(* PLC project LFAM, CODESYS CODESYS V3.5 SP22 Patch 4 *)
(* stored: creationDateTime 2026-11-11T00:00:00, modificationDateTime 2026-11-11T00:00:00 *)

PROGRAM PLC_PRG
  VAR
    PT_FUNDIDO_MPA : REAL;
    PT_FUNDIDO_RAW : INT;
    TT_SUBSTRATO_C : REAL;
    TT_SUBSTRATO_RAW : INT;
    TT_Z1 : REAL;
    TT_Z1_RAW : INT;
    TC_Z1_ABERTO : BOOL;
    TT_Z2 : REAL;
    TT_Z2_RAW : INT;
    TC_Z2_ABERTO : BOOL;
    TT_Z3 : REAL;
    TT_Z3_RAW : INT;
    TC_Z3_ABERTO : BOOL;
    TT_Z4 : REAL;
    TT_Z4_RAW : INT;
    TC_Z4_ABERTO : BOOL;
    TT_Z5 : REAL;
    TT_Z5_RAW : INT;
    TC_Z5_ABERTO : BOOL;
    TC_Z1_OK : BOOL;
    TC_Z2_OK : BOOL;
    TC_Z3_OK : BOOL;
    TC_Z4_OK : BOOL;
    TC_Z5_OK : BOOL;
    PLC_HEARTBEAT : INT;
    PWM_FASE : INT;
    PID_Z1 : Util.PID;
    SP_Z1 : REAL;
    Y_Z1 : REAL;
    LIM_Z1 : BOOL;
    OVF_Z1 : BOOL;
    PID_Z2 : Util.PID;
    SP_Z2 : REAL;
    Y_Z2 : REAL;
    LIM_Z2 : BOOL;
    OVF_Z2 : BOOL;
    PID_Z3 : Util.PID;
    SP_Z3 : REAL;
    Y_Z3 : REAL;
    LIM_Z3 : BOOL;
    OVF_Z3 : BOOL;
    PID_Z4 : Util.PID;
    SP_Z4 : REAL;
    Y_Z4 : REAL;
    LIM_Z4 : BOOL;
    OVF_Z4 : BOOL;
    PID_Z5 : Util.PID;
    SP_Z5 : REAL;
    Y_Z5 : REAL;
    LIM_Z5 : BOOL;
    OVF_Z5 : BOOL;
    PWM_Z1 : BOOL;
    PWM_Z2 : BOOL;
    PWM_Z3 : BOOL;
    PWM_Z4 : BOOL;
    PWM_Z5 : BOOL;
    PID_IR : Util.PID;
    SP_IR_C : REAL;
    Y_IR : REAL;
    LIM_IR : BOOL;
    OVF_IR : BOOL;
    PWM_IR : BOOL;
    SOBRETEMP_390_Z1 : BOOL;
    SOBRETEMP_390_Z2 : BOOL;
    SOBRETEMP_390_Z3 : BOOL;
    SOBRETEMP_390_Z4 : BOOL;
    SOBRETEMP_390_Z5 : BOOL;
    SOBRETEMP_400_Z1 : BOOL;
    SOBRETEMP_400_Z2 : BOOL;
    SOBRETEMP_400_Z3 : BOOL;
    SOBRETEMP_400_Z4 : BOOL;
    SOBRETEMP_400_Z5 : BOOL;
    SOBRETEMP_400 : BOOL;
    TC_FAULT : BOOL;
    TT_RESF : REAL;
    RESF_ACIMA_100 : BOOL;
    T_RESF_100C : TON;
    FALHA_RESF_2M : BOOL;
    EST_EXTRUSAO : BOOL;
    FUNIL_BAIXO : BOOL;
    ALIM_FUNIL : BOOL;
    T_FUNIL_VAZIO : TON;
    FALHA_SEM_MAT : BOOL;
    INV_RUN : BOOL;
    VENT_OK : BOOL;
    T_FALHA_VENT : TON;
    FALHA_VENT_10S : BOOL;
    K1_AQUEC : BOOL;
    K1_CONF : BOOL;
    T_K1_COLADO : TON;
    FALHA_K1_COL : BOOL;
    RESF_HI : BOOL;
    RESF_LO : BOOL;
    ALM_PRESSAO_16_5 : BOOL;
    PRESSAO_ALTA_17 : BOOL;
    SEG_OK : BOOL;
    MOT_SOBRETEMP : BOOL;
    INV_FALHA : BOOL;
    M_CAUSA : BOOL;
    FALHA_GERAL : BOOL;
    CAUSA_SEG_OK : BOOL;
    CAUSA_MOT_SOBRETEMP : BOOL;
    CAUSA_INV_FALHA : BOOL;
    CAUSA_PRESSAO_ALTA_17 : BOOL;
    CAUSA_SOBRETEMP_400 : BOOL;
    CAUSA_TC_FAULT : BOOL;
    CAUSA_FALHA_RESF_2M : BOOL;
    CAUSA_FALHA_SEM_MAT : BOOL;
    CAUSA_FALHA_VENT_10S : BOOL;
    CAUSA_FALHA_K1_COL : BOOL;
    BT_RESET : BOOL;
    BT_AQUEC : BOOL;
    EST_AQUEC : BOOL;
    DISJ_AQUEC : BOOL;
    RESF_ON : BOOL;
    Z1_ATEMP : BOOL;
    Z2_ATEMP : BOOL;
    Z3_ATEMP : BOOL;
    Z4_ATEMP : BOOL;
    Z5_ATEMP : BOOL;
    EST_ENCHARQUE : BOOL;
    T_ENCHARQUE : TON;
    ENCH_OK : BOOL;
    SECADOR_OK : BOOL;
    INV_PRONTO : BOOL;
    EST_PRONTO : BOOL;
    ROBO_EXT_PRONTA : BOOL;
    BT_DESLIGA : BOOL;
    SEL_AUTO : BOOL;
    BT_LIGA : BOOL;
    ROBO_CMD_EXTR : BOOL;
    VENT_MOTOR : BOOL;
    T_POS_VENT : TON;
    VENT_FIM : BOOL;
    REF_RPM_LIM : REAL;
    SP_RPM_OPERADOR : REAL;
    INV_REF : INT;
    SSR_Z1 : BOOL;
    SSR_Z2 : BOOL;
    SSR_Z3 : BOOL;
    SSR_Z4 : BOOL;
    SSR_Z5 : BOOL;
    IR_ACIMA_MIN : BOOL;
    IR_ABAIXO_MAX : BOOL;
    ROBO_EM_MOV : BOOL;
    IR_HAB : BOOL;
    SSR_IR : BOOL;
    TT_ZSR : REAL;
    ZSR_ABAIXO : BOOL;
    ALM_ZSR_BAIXA : BOOL;
    LUZ_VERDE : BOOL;
    LUZ_AMARELA : BOOL;
    LUZ_VERM_SIRENE : BOOL;
    RT_FUNIL : R_TRIG;
    FUNIL_PULSO : BOOL;
    CTU_LOTES : CTU;
    HMI_RESET_LOTES : BOOL;
    CONT_LOTES : WORD;
  END_VAR

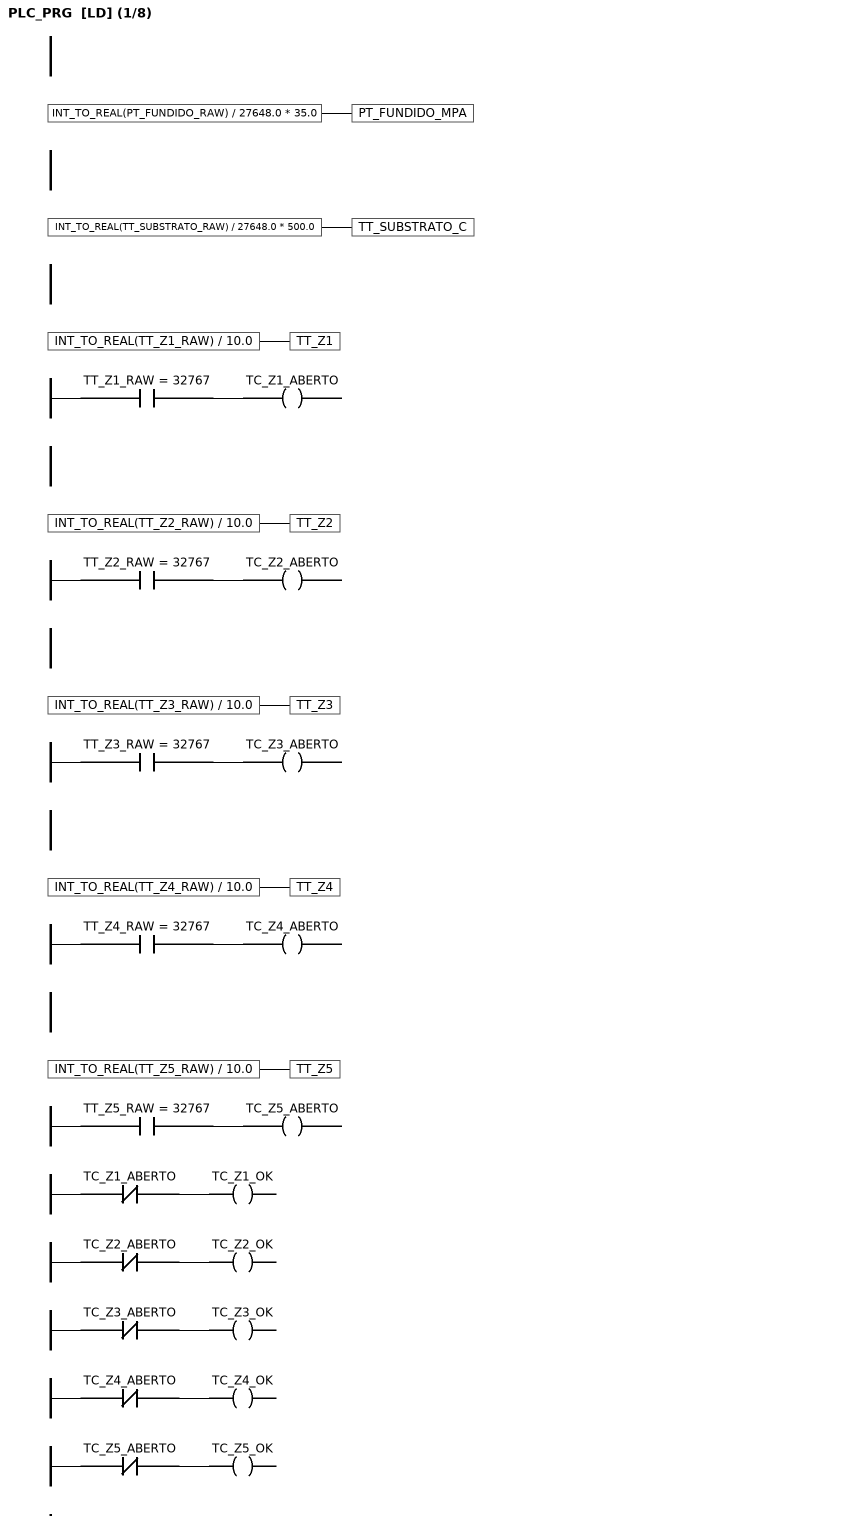
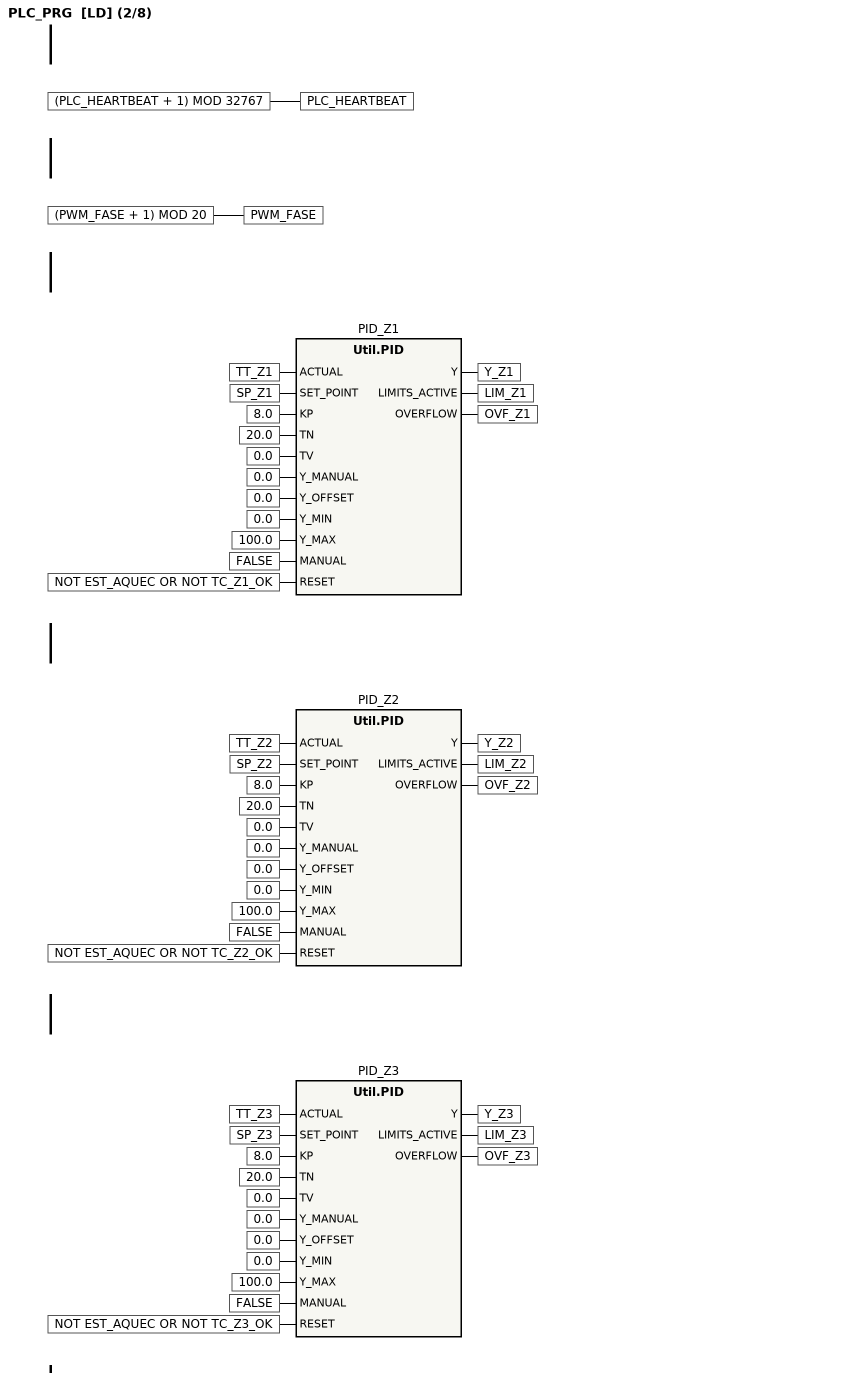
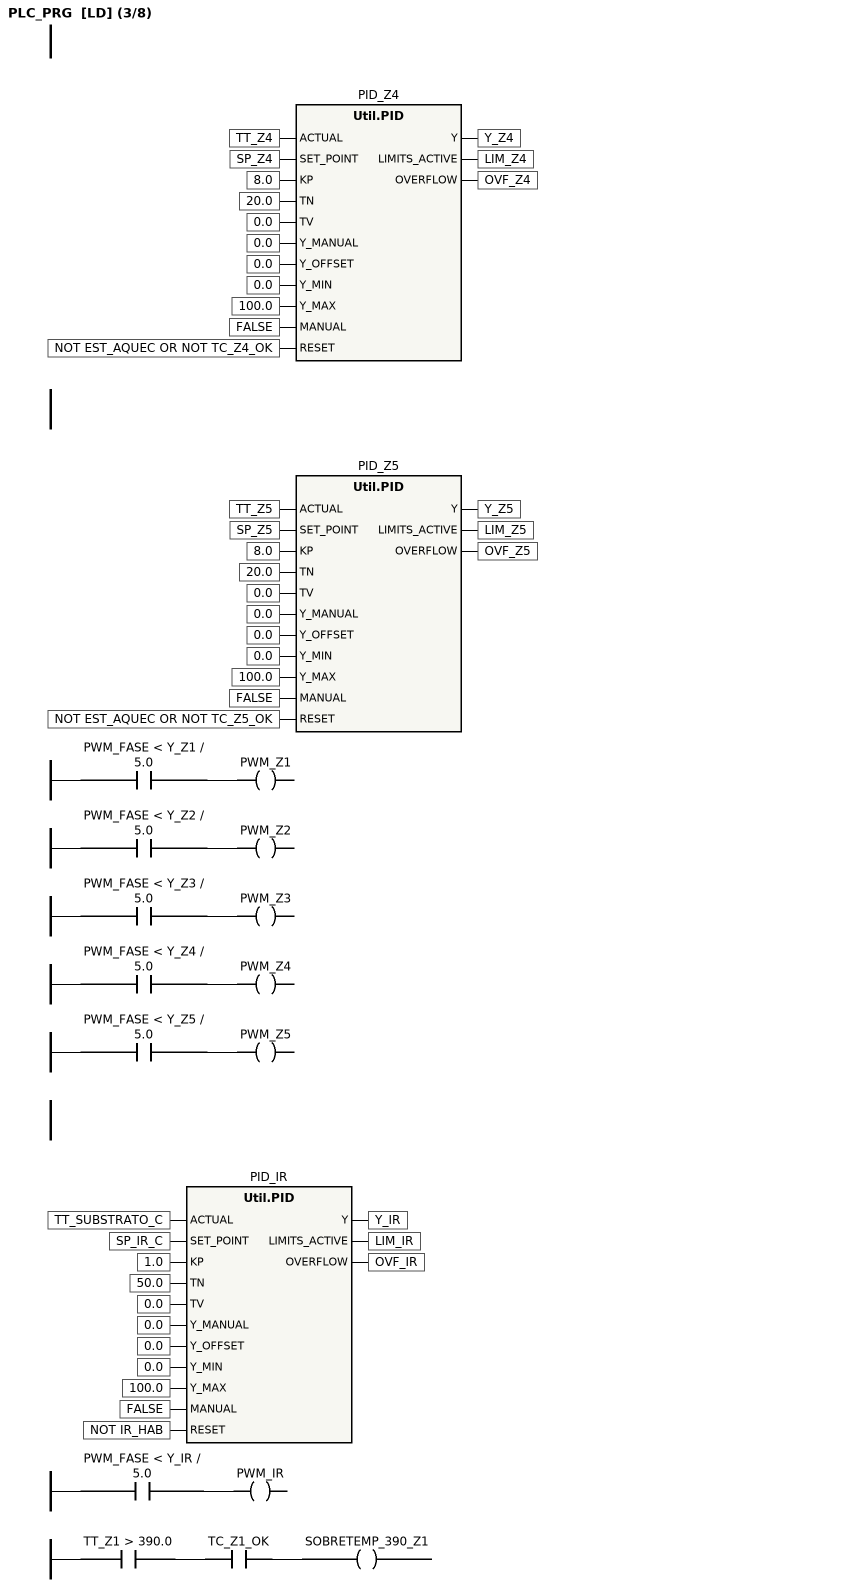
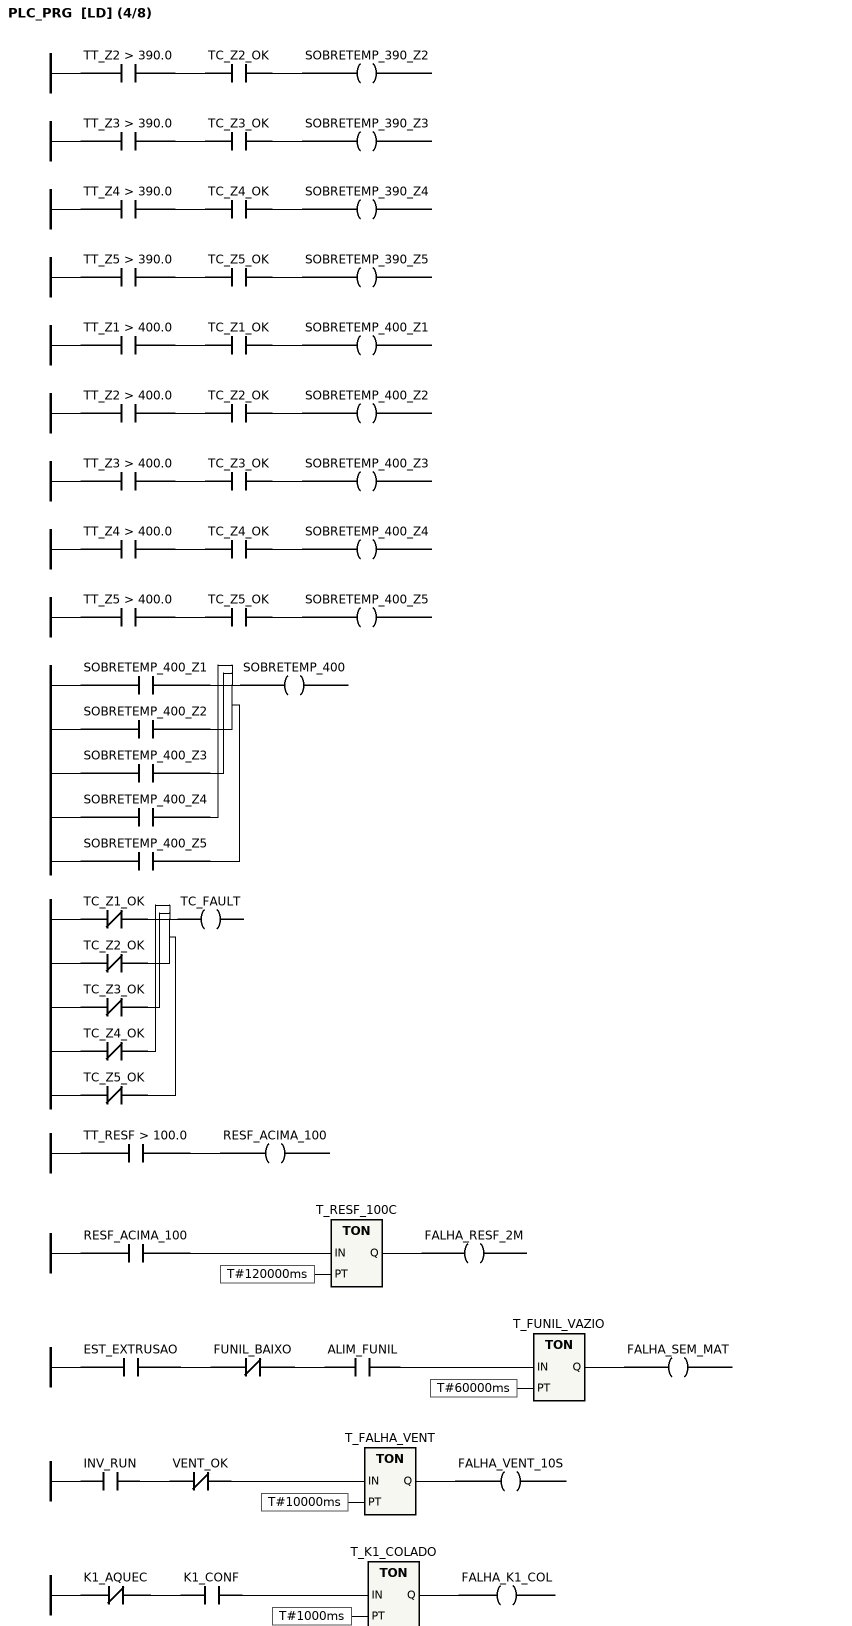
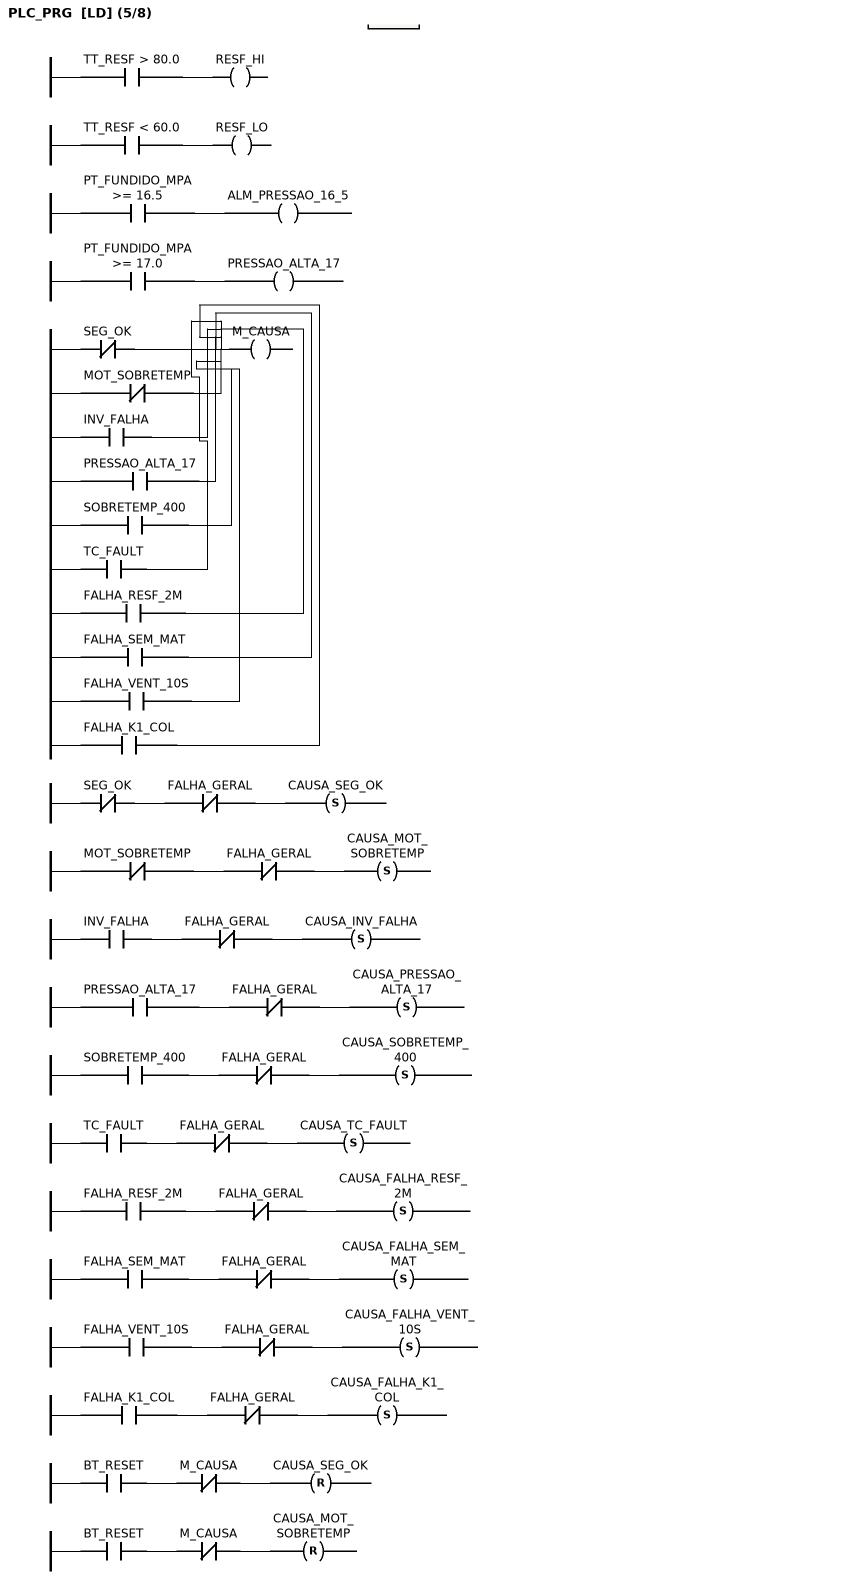
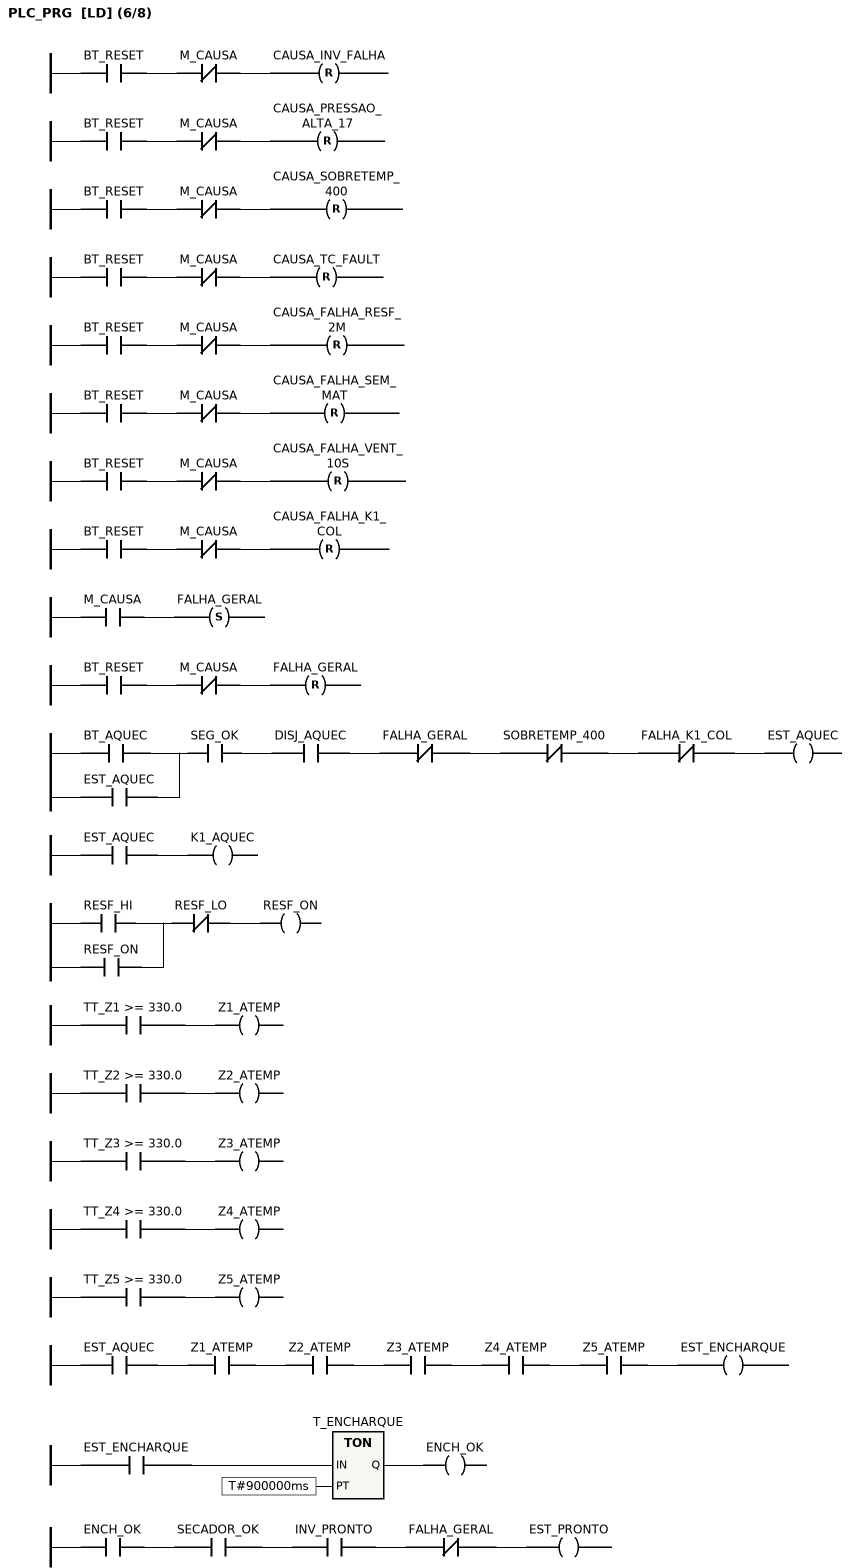
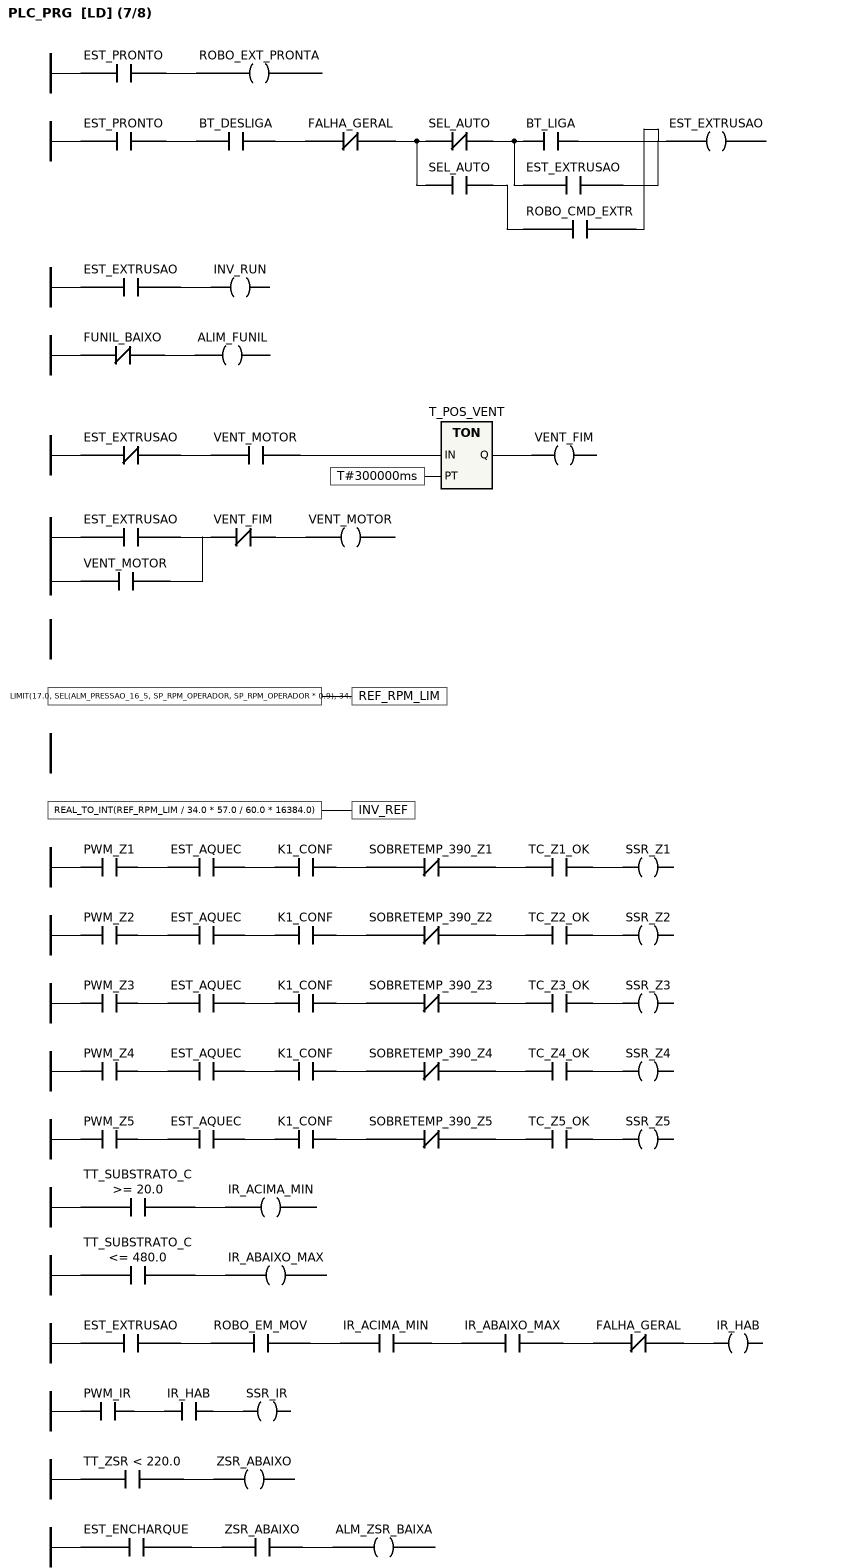
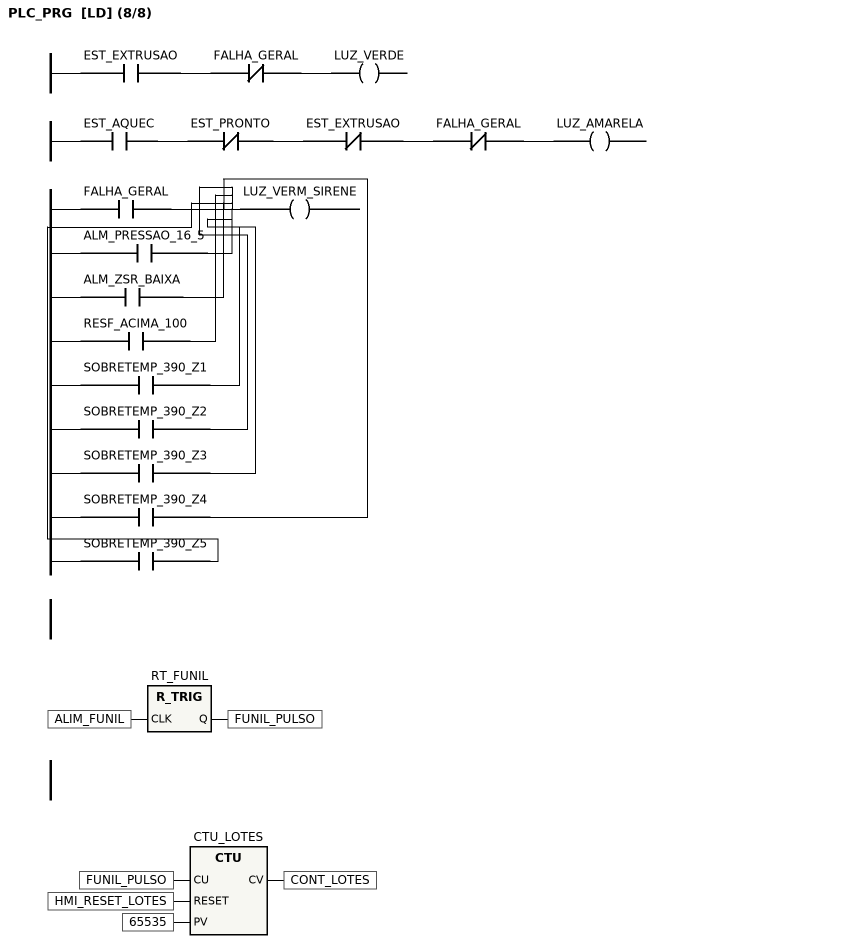
(* LD diagram, written out as Structured Text *)
(* NETWORK 01 - PT_FUNDIDO 0..27648 -> 0..35 MPa *)
PT_FUNDIDO_MPA := INT_TO_REAL(PT_FUNDIDO_RAW) / 27648.0 * 35.0;
(* NETWORK 01 - TT_SUBSTRATO 0..27648 -> 0..500 degC *)
TT_SUBSTRATO_C := INT_TO_REAL(TT_SUBSTRATO_RAW) / 27648.0 * 500.0;
(* NETWORK 02 - TT_Z1 (0,1 degC -> degC) *)
TT_Z1 := INT_TO_REAL(TT_Z1_RAW) / 10.0;
(* NETWORK 02 - Z1 termopar aberto (RAW = 32767) *)
TC_Z1_ABERTO := TT_Z1_RAW = 32767;
(* NETWORK 02 - TT_Z2 (0,1 degC -> degC) *)
TT_Z2 := INT_TO_REAL(TT_Z2_RAW) / 10.0;
(* NETWORK 02 - Z2 termopar aberto (RAW = 32767) *)
TC_Z2_ABERTO := TT_Z2_RAW = 32767;
(* NETWORK 02 - TT_Z3 (0,1 degC -> degC) *)
TT_Z3 := INT_TO_REAL(TT_Z3_RAW) / 10.0;
(* NETWORK 02 - Z3 termopar aberto (RAW = 32767) *)
TC_Z3_ABERTO := TT_Z3_RAW = 32767;
(* NETWORK 02 - TT_Z4 (0,1 degC -> degC) *)
TT_Z4 := INT_TO_REAL(TT_Z4_RAW) / 10.0;
(* NETWORK 02 - Z4 termopar aberto (RAW = 32767) *)
TC_Z4_ABERTO := TT_Z4_RAW = 32767;
(* NETWORK 02 - TT_Z5 (0,1 degC -> degC) *)
TT_Z5 := INT_TO_REAL(TT_Z5_RAW) / 10.0;
(* NETWORK 02 - Z5 termopar aberto (RAW = 32767) *)
TC_Z5_ABERTO := TT_Z5_RAW = 32767;
(* NETWORK 02 - TC_Z1_OK = nao aberto *)
TC_Z1_OK := NOT TC_Z1_ABERTO;
(* NETWORK 02 - TC_Z2_OK = nao aberto *)
TC_Z2_OK := NOT TC_Z2_ABERTO;
(* NETWORK 02 - TC_Z3_OK = nao aberto *)
TC_Z3_OK := NOT TC_Z3_ABERTO;
(* NETWORK 02 - TC_Z4_OK = nao aberto *)
TC_Z4_OK := NOT TC_Z4_ABERTO;
(* NETWORK 02 - TC_Z5_OK = nao aberto *)
TC_Z5_OK := NOT TC_Z5_ABERTO;
(* NETWORK 00 - PLC_HEARTBEAT: contador de vida do programa (INT, 0..32767) *)
PLC_HEARTBEAT := (PLC_HEARTBEAT + 1) MOD 32767;
(* NETWORK 06 - fase do PWM: (fase + 1) MOD 20 ciclos de 100 ms *)
PWM_FASE := (PWM_FASE + 1) MOD 20;
(* NETWORK 06 - PID zona 1 (Util.PID; RESET quando sem aquecimento ou termopar ruim) *)
PID_Z1(ACTUAL := TT_Z1, SET_POINT := SP_Z1, KP := 8.0, TN := 20.0, TV := 0.0, Y_MANUAL := 0.0, Y_OFFSET := 0.0, Y_MIN := 0.0, Y_MAX := 100.0, MANUAL := FALSE, RESET := NOT EST_AQUEC OR NOT TC_Z1_OK, Y => Y_Z1, LIMITS_ACTIVE => LIM_Z1, OVERFLOW => OVF_Z1);
(* NETWORK 06 - PID zona 2 (Util.PID; RESET quando sem aquecimento ou termopar ruim) *)
PID_Z2(ACTUAL := TT_Z2, SET_POINT := SP_Z2, KP := 8.0, TN := 20.0, TV := 0.0, Y_MANUAL := 0.0, Y_OFFSET := 0.0, Y_MIN := 0.0, Y_MAX := 100.0, MANUAL := FALSE, RESET := NOT EST_AQUEC OR NOT TC_Z2_OK, Y => Y_Z2, LIMITS_ACTIVE => LIM_Z2, OVERFLOW => OVF_Z2);
(* NETWORK 06 - PID zona 3 (Util.PID; RESET quando sem aquecimento ou termopar ruim) *)
PID_Z3(ACTUAL := TT_Z3, SET_POINT := SP_Z3, KP := 8.0, TN := 20.0, TV := 0.0, Y_MANUAL := 0.0, Y_OFFSET := 0.0, Y_MIN := 0.0, Y_MAX := 100.0, MANUAL := FALSE, RESET := NOT EST_AQUEC OR NOT TC_Z3_OK, Y => Y_Z3, LIMITS_ACTIVE => LIM_Z3, OVERFLOW => OVF_Z3);
(* NETWORK 06 - PID zona 4 (Util.PID; RESET quando sem aquecimento ou termopar ruim) *)
PID_Z4(ACTUAL := TT_Z4, SET_POINT := SP_Z4, KP := 8.0, TN := 20.0, TV := 0.0, Y_MANUAL := 0.0, Y_OFFSET := 0.0, Y_MIN := 0.0, Y_MAX := 100.0, MANUAL := FALSE, RESET := NOT EST_AQUEC OR NOT TC_Z4_OK, Y => Y_Z4, LIMITS_ACTIVE => LIM_Z4, OVERFLOW => OVF_Z4);
(* NETWORK 06 - PID zona 5 (Util.PID; RESET quando sem aquecimento ou termopar ruim) *)
PID_Z5(ACTUAL := TT_Z5, SET_POINT := SP_Z5, KP := 8.0, TN := 20.0, TV := 0.0, Y_MANUAL := 0.0, Y_OFFSET := 0.0, Y_MIN := 0.0, Y_MAX := 100.0, MANUAL := FALSE, RESET := NOT EST_AQUEC OR NOT TC_Z5_OK, Y => Y_Z5, LIMITS_ACTIVE => LIM_Z5, OVERFLOW => OVF_Z5);
(* NETWORK 06 - PWM_Z1: fase < saida do PID (% x 20 ciclos) *)
PWM_Z1 := PWM_FASE < Y_Z1 / 5.0;
(* NETWORK 06 - PWM_Z2: fase < saida do PID (% x 20 ciclos) *)
PWM_Z2 := PWM_FASE < Y_Z2 / 5.0;
(* NETWORK 06 - PWM_Z3: fase < saida do PID (% x 20 ciclos) *)
PWM_Z3 := PWM_FASE < Y_Z3 / 5.0;
(* NETWORK 06 - PWM_Z4: fase < saida do PID (% x 20 ciclos) *)
PWM_Z4 := PWM_FASE < Y_Z4 / 5.0;
(* NETWORK 06 - PWM_Z5: fase < saida do PID (% x 20 ciclos) *)
PWM_Z5 := PWM_FASE < Y_Z5 / 5.0;
(* NETWORK 13 - PID do aquecedor IR (RESET quando IR nao habilitado) *)
PID_IR(ACTUAL := TT_SUBSTRATO_C, SET_POINT := SP_IR_C, KP := 1.0, TN := 50.0, TV := 0.0, Y_MANUAL := 0.0, Y_OFFSET := 0.0, Y_MIN := 0.0, Y_MAX := 100.0, MANUAL := FALSE, RESET := NOT IR_HAB, Y => Y_IR, LIMITS_ACTIVE => LIM_IR, OVERFLOW => OVF_IR);
(* NETWORK 13 - PWM_IR: fase < saida do PID (% x 20 ciclos) *)
PWM_IR := PWM_FASE < Y_IR / 5.0;
(* NETWORK 02 - Z1 acima de 390 degC (pre-alarme; so com termopar valido) *)
SOBRETEMP_390_Z1 := (TT_Z1 > 390.0) AND TC_Z1_OK;
(* NETWORK 02 - Z2 acima de 390 degC (pre-alarme; so com termopar valido) *)
SOBRETEMP_390_Z2 := (TT_Z2 > 390.0) AND TC_Z2_OK;
(* NETWORK 02 - Z3 acima de 390 degC (pre-alarme; so com termopar valido) *)
SOBRETEMP_390_Z3 := (TT_Z3 > 390.0) AND TC_Z3_OK;
(* NETWORK 02 - Z4 acima de 390 degC (pre-alarme; so com termopar valido) *)
SOBRETEMP_390_Z4 := (TT_Z4 > 390.0) AND TC_Z4_OK;
(* NETWORK 02 - Z5 acima de 390 degC (pre-alarme; so com termopar valido) *)
SOBRETEMP_390_Z5 := (TT_Z5 > 390.0) AND TC_Z5_OK;
(* NETWORK 02 - Z1 acima de 400 degC (falha; so com termopar valido: fio aberto le 3276,7 e NAO e sobretemperatura) *)
SOBRETEMP_400_Z1 := (TT_Z1 > 400.0) AND TC_Z1_OK;
(* NETWORK 02 - Z2 acima de 400 degC (falha; so com termopar valido: fio aberto le 3276,7 e NAO e sobretemperatura) *)
SOBRETEMP_400_Z2 := (TT_Z2 > 400.0) AND TC_Z2_OK;
(* NETWORK 02 - Z3 acima de 400 degC (falha; so com termopar valido: fio aberto le 3276,7 e NAO e sobretemperatura) *)
SOBRETEMP_400_Z3 := (TT_Z3 > 400.0) AND TC_Z3_OK;
(* NETWORK 02 - Z4 acima de 400 degC (falha; so com termopar valido: fio aberto le 3276,7 e NAO e sobretemperatura) *)
SOBRETEMP_400_Z4 := (TT_Z4 > 400.0) AND TC_Z4_OK;
(* NETWORK 02 - Z5 acima de 400 degC (falha; so com termopar valido: fio aberto le 3276,7 e NAO e sobretemperatura) *)
SOBRETEMP_400_Z5 := (TT_Z5 > 400.0) AND TC_Z5_OK;
(* NETWORK 02 - SOBRETEMP_400: OR das cinco zonas *)
SOBRETEMP_400 := SOBRETEMP_400_Z1 OR SOBRETEMP_400_Z2 OR SOBRETEMP_400_Z3 OR SOBRETEMP_400_Z4 OR SOBRETEMP_400_Z5;
(* NETWORK 02 - TC_FAULT: OR de termopar com qualidade ruim *)
TC_FAULT := NOT TC_Z1_OK OR NOT TC_Z2_OK OR NOT TC_Z3_OK OR NOT TC_Z4_OK OR NOT TC_Z5_OK;
(* NETWORK 03 - TT_RESF acima de 100 degC *)
RESF_ACIMA_100 := TT_RESF > 100.0;
(* NETWORK 03 - camara quente por 2 min *)
T_RESF_100C(IN := RESF_ACIMA_100, PT := T#120000ms);
FALHA_RESF_2M := T_RESF_100C.Q;
(* NETWORK 03 - sem material por 60 s (FUNIL_BAIXO=0 e vazio) *)
T_FUNIL_VAZIO(IN := EST_EXTRUSAO AND NOT FUNIL_BAIXO AND ALIM_FUNIL, PT := T#60000ms);
FALHA_SEM_MAT := T_FUNIL_VAZIO.Q;
(* NETWORK 03 - rosca sem ventilacao por 10 s *)
T_FALHA_VENT(IN := INV_RUN AND NOT VENT_OK, PT := T#10000ms);
FALHA_VENT_10S := T_FALHA_VENT.Q;
(* NETWORK 03 - K1 colado por 1 s (confirma sem comando) *)
T_K1_COLADO(IN := NOT K1_AQUEC AND K1_CONF, PT := T#1000ms);
FALHA_K1_COL := T_K1_COLADO.Q;
(* NETWORK 07 - RESF_HI: TT_RESF acima de 80 degC *)
RESF_HI := TT_RESF > 80.0;
(* NETWORK 07 - RESF_LO: TT_RESF abaixo de 60 degC *)
RESF_LO := TT_RESF < 60.0;
(* NETWORK 12 - ALM_PRESSAO_16_5: pressao >= 16,5 MPa *)
ALM_PRESSAO_16_5 := PT_FUNDIDO_MPA >= 16.5;
(* NETWORK 04 - PRESSAO_ALTA_17: pressao >= 17 MPa *)
PRESSAO_ALTA_17 := PT_FUNDIDO_MPA >= 17.0;
(* NETWORK 04a - M_CAUSA: OR de todas as causas criticas *)
M_CAUSA := NOT SEG_OK OR NOT MOT_SOBRETEMP OR INV_FALHA OR PRESSAO_ALTA_17 OR SOBRETEMP_400 OR TC_FAULT OR FALHA_RESF_2M OR FALHA_SEM_MAT OR FALHA_VENT_10S OR FALHA_K1_COL;
(* NETWORK 04d - primeira causa: CAUSA_SEG_OK (set na varredura em que a falha ainda nao estava travada) *)
IF NOT SEG_OK AND NOT FALHA_GERAL THEN CAUSA_SEG_OK := TRUE; END_IF;
(* NETWORK 04d - primeira causa: CAUSA_MOT_SOBRETEMP (set na varredura em que a falha ainda nao estava travada) *)
IF NOT MOT_SOBRETEMP AND NOT FALHA_GERAL THEN CAUSA_MOT_SOBRETEMP := TRUE; END_IF;
(* NETWORK 04d - primeira causa: CAUSA_INV_FALHA (set na varredura em que a falha ainda nao estava travada) *)
IF INV_FALHA AND NOT FALHA_GERAL THEN CAUSA_INV_FALHA := TRUE; END_IF;
(* NETWORK 04d - primeira causa: CAUSA_PRESSAO_ALTA_17 (set na varredura em que a falha ainda nao estava travada) *)
IF PRESSAO_ALTA_17 AND NOT FALHA_GERAL THEN CAUSA_PRESSAO_ALTA_17 := TRUE; END_IF;
(* NETWORK 04d - primeira causa: CAUSA_SOBRETEMP_400 (set na varredura em que a falha ainda nao estava travada) *)
IF SOBRETEMP_400 AND NOT FALHA_GERAL THEN CAUSA_SOBRETEMP_400 := TRUE; END_IF;
(* NETWORK 04d - primeira causa: CAUSA_TC_FAULT (set na varredura em que a falha ainda nao estava travada) *)
IF TC_FAULT AND NOT FALHA_GERAL THEN CAUSA_TC_FAULT := TRUE; END_IF;
(* NETWORK 04d - primeira causa: CAUSA_FALHA_RESF_2M (set na varredura em que a falha ainda nao estava travada) *)
IF FALHA_RESF_2M AND NOT FALHA_GERAL THEN CAUSA_FALHA_RESF_2M := TRUE; END_IF;
(* NETWORK 04d - primeira causa: CAUSA_FALHA_SEM_MAT (set na varredura em que a falha ainda nao estava travada) *)
IF FALHA_SEM_MAT AND NOT FALHA_GERAL THEN CAUSA_FALHA_SEM_MAT := TRUE; END_IF;
(* NETWORK 04d - primeira causa: CAUSA_FALHA_VENT_10S (set na varredura em que a falha ainda nao estava travada) *)
IF FALHA_VENT_10S AND NOT FALHA_GERAL THEN CAUSA_FALHA_VENT_10S := TRUE; END_IF;
(* NETWORK 04d - primeira causa: CAUSA_FALHA_K1_COL (set na varredura em que a falha ainda nao estava travada) *)
IF FALHA_K1_COL AND NOT FALHA_GERAL THEN CAUSA_FALHA_K1_COL := TRUE; END_IF;
(* NETWORK 04e - CAUSA_SEG_OK reseta junto com a falha (BT_RESET e nenhuma causa ativa) *)
IF BT_RESET AND NOT M_CAUSA THEN CAUSA_SEG_OK := FALSE; END_IF;
(* NETWORK 04e - CAUSA_MOT_SOBRETEMP reseta junto com a falha (BT_RESET e nenhuma causa ativa) *)
IF BT_RESET AND NOT M_CAUSA THEN CAUSA_MOT_SOBRETEMP := FALSE; END_IF;
(* NETWORK 04e - CAUSA_INV_FALHA reseta junto com a falha (BT_RESET e nenhuma causa ativa) *)
IF BT_RESET AND NOT M_CAUSA THEN CAUSA_INV_FALHA := FALSE; END_IF;
(* NETWORK 04e - CAUSA_PRESSAO_ALTA_17 reseta junto com a falha (BT_RESET e nenhuma causa ativa) *)
IF BT_RESET AND NOT M_CAUSA THEN CAUSA_PRESSAO_ALTA_17 := FALSE; END_IF;
(* NETWORK 04e - CAUSA_SOBRETEMP_400 reseta junto com a falha (BT_RESET e nenhuma causa ativa) *)
IF BT_RESET AND NOT M_CAUSA THEN CAUSA_SOBRETEMP_400 := FALSE; END_IF;
(* NETWORK 04e - CAUSA_TC_FAULT reseta junto com a falha (BT_RESET e nenhuma causa ativa) *)
IF BT_RESET AND NOT M_CAUSA THEN CAUSA_TC_FAULT := FALSE; END_IF;
(* NETWORK 04e - CAUSA_FALHA_RESF_2M reseta junto com a falha (BT_RESET e nenhuma causa ativa) *)
IF BT_RESET AND NOT M_CAUSA THEN CAUSA_FALHA_RESF_2M := FALSE; END_IF;
(* NETWORK 04e - CAUSA_FALHA_SEM_MAT reseta junto com a falha (BT_RESET e nenhuma causa ativa) *)
IF BT_RESET AND NOT M_CAUSA THEN CAUSA_FALHA_SEM_MAT := FALSE; END_IF;
(* NETWORK 04e - CAUSA_FALHA_VENT_10S reseta junto com a falha (BT_RESET e nenhuma causa ativa) *)
IF BT_RESET AND NOT M_CAUSA THEN CAUSA_FALHA_VENT_10S := FALSE; END_IF;
(* NETWORK 04e - CAUSA_FALHA_K1_COL reseta junto com a falha (BT_RESET e nenhuma causa ativa) *)
IF BT_RESET AND NOT M_CAUSA THEN CAUSA_FALHA_K1_COL := FALSE; END_IF;
(* NETWORK 04b - FALHA_GERAL travada (SET por M_CAUSA) *)
IF M_CAUSA THEN FALHA_GERAL := TRUE; END_IF;
(* NETWORK 04c - RESET condicionado (BT_RESET e nenhuma causa ativa) *)
IF BT_RESET AND NOT M_CAUSA THEN FALHA_GERAL := FALSE; END_IF;
(* NETWORK 05 - EST_AQUEC (selo; desligamento tem prioridade) *)
EST_AQUEC := (BT_AQUEC OR EST_AQUEC) AND SEG_OK AND DISJ_AQUEC AND NOT FALHA_GERAL AND NOT SOBRETEMP_400 AND NOT FALHA_K1_COL;
(* NETWORK 05b - K1_AQUEC segue EST_AQUEC (unico escritor) *)
K1_AQUEC := EST_AQUEC;
(* NETWORK 07 - Resfriamento por histerese (liga >80, mantem ate <60) *)
RESF_ON := (RESF_HI OR RESF_ON) AND NOT RESF_LO;
(* NETWORK 08 - Z1 >= 330 degC *)
Z1_ATEMP := TT_Z1 >= 330.0;
(* NETWORK 08 - Z2 >= 330 degC *)
Z2_ATEMP := TT_Z2 >= 330.0;
(* NETWORK 08 - Z3 >= 330 degC *)
Z3_ATEMP := TT_Z3 >= 330.0;
(* NETWORK 08 - Z4 >= 330 degC *)
Z4_ATEMP := TT_Z4 >= 330.0;
(* NETWORK 08 - Z5 >= 330 degC *)
Z5_ATEMP := TT_Z5 >= 330.0;
(* NETWORK 08 - EST_ENCHARQUE: aquecimento ligado e todas as zonas >= 330 (Prancha 2: gate por EST_AQUEC) *)
EST_ENCHARQUE := EST_AQUEC AND Z1_ATEMP AND Z2_ATEMP AND Z3_ATEMP AND Z4_ATEMP AND Z5_ATEMP;
(* NETWORK 08 - encharque continuo de 15 min *)
T_ENCHARQUE(IN := EST_ENCHARQUE, PT := T#900000ms);
ENCH_OK := T_ENCHARQUE.Q;
(* NETWORK 09 - EST_PRONTO: encharque ok, secador, inversor pronto, sem falha memorizada *)
EST_PRONTO := ENCH_OK AND SECADOR_OK AND INV_PRONTO AND NOT FALHA_GERAL;
(* NETWORK 09 - ROBO_EXT_PRONTA segue EST_PRONTO *)
ROBO_EXT_PRONTA := EST_PRONTO;
(* NETWORK 10 - Rosca (manual com selo / automatico pelo robo) *)
EST_EXTRUSAO := EST_PRONTO AND BT_DESLIGA AND NOT FALHA_GERAL AND (NOT SEL_AUTO AND BT_LIGA OR NOT SEL_AUTO AND EST_EXTRUSAO OR SEL_AUTO AND ROBO_CMD_EXTR);
(* NETWORK 10 - INV_RUN segue EST_EXTRUSAO (unico escritor) *)
INV_RUN := EST_EXTRUSAO;
(* NETWORK 14 - ALIM_FUNIL: carregador liga com funil vazio (FUNIL_BAIXO=0) *)
ALIM_FUNIL := NOT FUNIL_BAIXO;
(* NETWORK 11 - 5 min de pos-ventilacao (rosca parada e ventilador ligado) *)
T_POS_VENT(IN := NOT EST_EXTRUSAO AND VENT_MOTOR, PT := T#300000ms);
VENT_FIM := T_POS_VENT.Q;
(* NETWORK 11 - VENT_MOTOR (unico escritor): rosca OU em pos-ventilacao ate o fim do tempo *)
VENT_MOTOR := (EST_EXTRUSAO OR VENT_MOTOR) AND NOT VENT_FIM;
(* NETWORK 12 - REF_RPM_LIM := LIMIT(17, SP (x0,9 se alarme), 34) - unico escritor *)
REF_RPM_LIM := LIMIT(17.0, SEL(ALM_PRESSAO_16_5, SP_RPM_OPERADOR, SP_RPM_OPERADOR * 0.9), 34.0);
(* NETWORK 12 - INV_REF (unico escritor): rpm -> escala do inversor (hipotese 16384 = 60 Hz) *)
INV_REF := REAL_TO_INT(REF_RPM_LIM / 34.0 * 57.0 / 60.0 * 16384.0);
(* NETWORK 06 - SSR_Z1: PWM so com aquecimento, K1 confirmado, zona < 390 degC e termopar integro *)
SSR_Z1 := PWM_Z1 AND EST_AQUEC AND K1_CONF AND NOT SOBRETEMP_390_Z1 AND TC_Z1_OK;
(* NETWORK 06 - SSR_Z2: PWM so com aquecimento, K1 confirmado, zona < 390 degC e termopar integro *)
SSR_Z2 := PWM_Z2 AND EST_AQUEC AND K1_CONF AND NOT SOBRETEMP_390_Z2 AND TC_Z2_OK;
(* NETWORK 06 - SSR_Z3: PWM so com aquecimento, K1 confirmado, zona < 390 degC e termopar integro *)
SSR_Z3 := PWM_Z3 AND EST_AQUEC AND K1_CONF AND NOT SOBRETEMP_390_Z3 AND TC_Z3_OK;
(* NETWORK 06 - SSR_Z4: PWM so com aquecimento, K1 confirmado, zona < 390 degC e termopar integro *)
SSR_Z4 := PWM_Z4 AND EST_AQUEC AND K1_CONF AND NOT SOBRETEMP_390_Z4 AND TC_Z4_OK;
(* NETWORK 06 - SSR_Z5: PWM so com aquecimento, K1 confirmado, zona < 390 degC e termopar integro *)
SSR_Z5 := PWM_Z5 AND EST_AQUEC AND K1_CONF AND NOT SOBRETEMP_390_Z5 AND TC_Z5_OK;
(* NETWORK 13 - IR_FAIXA_MIN: substrato >= 20 degC *)
IR_ACIMA_MIN := TT_SUBSTRATO_C >= 20.0;
(* NETWORK 13 - IR_FAIXA_MAX: substrato <= 480 degC *)
IR_ABAIXO_MAX := TT_SUBSTRATO_C <= 480.0;
(* NETWORK 13 - IR_HAB: rosca girando, robo em movimento, pirometro na faixa, sem falha *)
IR_HAB := EST_EXTRUSAO AND ROBO_EM_MOV AND IR_ACIMA_MIN AND IR_ABAIXO_MAX AND NOT FALHA_GERAL;
(* NETWORK 13 - SSR_IR (unico escritor): PWM_IR so com IR_HAB *)
SSR_IR := PWM_IR AND IR_HAB;
(* NETWORK 15 - ZSR_ABAIXO: trecho sem resistencia < 220 degC *)
ZSR_ABAIXO := TT_ZSR < 220.0;
(* NETWORK 15 - ALM_ZSR_BAIXA: so durante o encharque (Prancha 4) *)
ALM_ZSR_BAIXA := EST_ENCHARQUE AND ZSR_ABAIXO;
(* NETWORK 15 - LUZ_VERDE: extrusao sem falha travada *)
LUZ_VERDE := EST_EXTRUSAO AND NOT FALHA_GERAL;
(* NETWORK 15 - LUZ_AMARELA: aquecendo ou aguardando encharque (nao pronto, sem extrusao, sem falha) *)
LUZ_AMARELA := EST_AQUEC AND NOT EST_PRONTO AND NOT EST_EXTRUSAO AND NOT FALHA_GERAL;
(* NETWORK 15 - LUZ_VERM_SIRENE: falha travada OU pressao 16,5 OU trecho frio OU zona > 390 OU camara > 100 degC *)
LUZ_VERM_SIRENE := FALHA_GERAL OR ALM_PRESSAO_16_5 OR ALM_ZSR_BAIXA OR RESF_ACIMA_100 OR SOBRETEMP_390_Z1 OR SOBRETEMP_390_Z2 OR SOBRETEMP_390_Z3 OR SOBRETEMP_390_Z4 OR SOBRETEMP_390_Z5;
(* NETWORK 14 - R_TRIG: borda de subida do carregador *)
RT_FUNIL(CLK := ALIM_FUNIL, Q => FUNIL_PULSO);
(* NETWORK 14 - CTU: recargas do dosador (reset pelo SCADA) *)
CTU_LOTES(CU := FUNIL_PULSO, RESET := HMI_RESET_LOTES, PV := 65535, CV => CONT_LOTES);
END_PROGRAM
